{region 'Documentation'}
(*!
<summary>Checks children already Completed at the first helper call after their Start.</summary>
*)
{endregion}
FUNCTION_BLOCK Test_SerialImmediateCompletion EXTENDS OrchestrationTestBase

SUPER^();

{region 'Documentation'}
(*!
<summary>Defines this scenario independently of the subject's internal fields.</summary>
*)
{endregion}
METHOD PROTECTED ConfigureScenario
FArrayLayout := E_OrchestrationArrayLayout.Ordinary;
FChildCount := 3;
FStepCount := 8;

{region "Cycle 01 - Idle readiness"}
FSteps[1].Task := E_OrchestratorTask.Idle;
FSteps[1].ExpectedReady := TRUE;
{endregion}

{region "Cycle 02 - Start child 1"}
FSteps[2].Children[1].State := E_State.Completed;
FSteps[2].Children[1].Ready := FALSE;
FSteps[2].Children[1].Complete := TRUE;
FSteps[2].Children[1].Result := E_Result.Passed;
FSteps[2].ExpectedStartChild := 1;
FSteps[2].ExpectedSlot := 1;
FSteps[2].ExpectedReservations[1] := 1;
{endregion}

{region "Cycle 03 - Reconcile completed child 1"}
FSteps[3].Children[1].State := E_State.Completed;
FSteps[3].Children[1].Ready := FALSE;
FSteps[3].Children[1].Complete := TRUE;
FSteps[3].Children[1].Result := E_Result.Passed;
FSteps[3].ExpectedSlot := 2;
FSteps[3].ExpectedReleasedEntries[1] := 1;
{endregion}

{region "Cycle 04 - Start child 2"}
FSteps[4].Children[1].State := E_State.Completed;
FSteps[4].Children[1].Ready := FALSE;
FSteps[4].Children[1].Complete := TRUE;
FSteps[4].Children[1].Result := E_Result.Passed;
FSteps[4].Children[2].State := E_State.Completed;
FSteps[4].Children[2].Ready := FALSE;
FSteps[4].Children[2].Complete := TRUE;
FSteps[4].Children[2].Result := E_Result.Passed;
FSteps[4].ExpectedStartChild := 2;
FSteps[4].ExpectedSlot := 2;
FSteps[4].ExpectedReservations[2] := 1;
{endregion}

{region "Cycle 05 - Reconcile completed child 2"}
FSteps[5].Children[1].State := E_State.Completed;
FSteps[5].Children[1].Ready := FALSE;
FSteps[5].Children[1].Complete := TRUE;
FSteps[5].Children[1].Result := E_Result.Passed;
FSteps[5].Children[2].State := E_State.Completed;
FSteps[5].Children[2].Ready := FALSE;
FSteps[5].Children[2].Complete := TRUE;
FSteps[5].Children[2].Result := E_Result.Passed;
FSteps[5].ExpectedSlot := 3;
FSteps[5].ExpectedReleasedEntries[2] := 1;
{endregion}

{region "Cycle 06 - Start child 3"}
FSteps[6].Children[1].State := E_State.Completed;
FSteps[6].Children[1].Ready := FALSE;
FSteps[6].Children[1].Complete := TRUE;
FSteps[6].Children[1].Result := E_Result.Passed;
FSteps[6].Children[2].State := E_State.Completed;
FSteps[6].Children[2].Ready := FALSE;
FSteps[6].Children[2].Complete := TRUE;
FSteps[6].Children[2].Result := E_Result.Passed;
FSteps[6].Children[3].State := E_State.Completed;
FSteps[6].Children[3].Ready := FALSE;
FSteps[6].Children[3].Complete := TRUE;
FSteps[6].Children[3].Result := E_Result.Passed;
FSteps[6].ExpectedStartChild := 3;
FSteps[6].ExpectedSlot := 3;
FSteps[6].ExpectedReservations[3] := 1;
{endregion}

{region "Cycle 07 - Completed observation"}
FSteps[7].Children[1].State := E_State.Completed;
FSteps[7].Children[1].Ready := FALSE;
FSteps[7].Children[1].Complete := TRUE;
FSteps[7].Children[1].Result := E_Result.Passed;
FSteps[7].Children[2].State := E_State.Completed;
FSteps[7].Children[2].Ready := FALSE;
FSteps[7].Children[2].Complete := TRUE;
FSteps[7].Children[2].Result := E_Result.Passed;
FSteps[7].Children[3].State := E_State.Completed;
FSteps[7].Children[3].Ready := FALSE;
FSteps[7].Children[3].Complete := TRUE;
FSteps[7].Children[3].Result := E_Result.Passed;
FSteps[7].ExpectedReleasedEntries[3] := 1;
FSteps[7].ExpectedFinished := TRUE;
{endregion}

{region "Cycle 08 - Completed observation"}
FSteps[8].Children[1].State := E_State.Completed;
FSteps[8].Children[1].Ready := FALSE;
FSteps[8].Children[1].Complete := TRUE;
FSteps[8].Children[1].Result := E_Result.Passed;
FSteps[8].Children[2].State := E_State.Completed;
FSteps[8].Children[2].Ready := FALSE;
FSteps[8].Children[2].Complete := TRUE;
FSteps[8].Children[2].Result := E_Result.Passed;
FSteps[8].Children[3].State := E_State.Completed;
FSteps[8].Children[3].Ready := FALSE;
FSteps[8].Children[3].Complete := TRUE;
FSteps[8].Children[3].Result := E_Result.Passed;
FSteps[8].ExpectedFinished := TRUE;
{endregion}
END_METHOD

END_FUNCTION_BLOCK

(* stored: Version 1.1.0.1
   POU Test_SerialImmediateCompletion: Id {fa36fb4b-4420-4cd5-92cc-ed7b9b008dc9}, SpecialFunc None
   Folder Internal: Id {5d46dc73-efa4-43b3-9347-7b7ebd89049e}
   Method ConfigureScenario: Id {0d4328a5-6b6a-42dc-89e4-eb9a57e7f97a} *)
